(* IEC 61131-3 sources: Lasal-MCP/examples/SampleSource/5_ClassInputOutputSolution/Stations/MachineControl/MachineControl/Class/AlarmStation, 1 file *)

(* ---- AlarmStation.st ---- *)
(*!
<Class
	Name               = "AlarmStation"
	Revision           = "1.2"
	RealtimeTask       = "false"
	CyclicTask         = "false"
	BackgroundTask     = "false"
	Sigmatek           = "true"
	OSInterface        = "false"
	HighPriority       = "false"
	Automatic          = "false"
	UpdateMode         = "Prescan"
	SharedCommandTable = "true"
	Objectsize         = "(586,120)"
	Comment            = "Class collected number of active op-mode alarms and delivers this informations to the class AlarmBufferBase.">
	<Channels>
		<Server Name="ClassSvr" Visualized="false" Initialize="false" WriteProtected="true" Retentive="false"/>
		<Client Name="Active" Required="false" Internal="false"/>
		<Client Name="AlarmInfo" Required="false" Internal="false"/>
		<Client Name="coAlarmBufferBase" Required="true" Internal="false"/>
		<Client Name="GroupAutomatic" Required="false" Internal="false"/>
		<Client Name="GroupError" Required="false" Internal="false"/>
		<Client Name="GroupHoming" Required="false" Internal="false"/>
		<Client Name="GroupInit" Required="false" Internal="false"/>
		<Client Name="GroupManual" Required="false" Internal="false"/>
		<Client Name="GroupSemiAuto" Required="false" Internal="false"/>
		<Client Name="GroupSetup" Required="false" Internal="false"/>
		<Client Name="GroupStop" Required="false" Internal="false"/>
	</Channels>
	<RevDoku>
		<Owner Company="Sigmatek" Author="ObeChr"/>
		<Dokumentation Revision="1.2" Date="2017-07-26" Author="KruAle" Company="Sigmatek" Description="Added client to deactivate class if station is not available."/>
		<Dokumentation Revision="1.1" Date="2016-08-09" Author="ObeChr" Company="Sigmatek" Description="Added client to get AlarmInfo from other stations."/>
		<Dokumentation Revision="1.0" Date="2016-03-23" Author="ObeChr" Company="Sigmatek" Description="First library version."/>
	</RevDoku>
</Class>
*)
AlarmStation : CLASS
  //Servers:
	ClassSvr 	: SvrChCmd_DINT;
  //Clients:
	coAlarmBufferBase 	: CltChCmd_AlarmBufferBase;
	Active 	: CltCh_DINT;
	GroupInit 	: CltCh_UDINT;
	GroupHoming 	: CltCh_UDINT;
	GroupStop 	: CltCh_UDINT;
	GroupSetup 	: CltCh_UDINT;
	GroupManual 	: CltCh_UDINT;
	GroupSemiAuto 	: CltCh_UDINT;
	GroupAutomatic 	: CltCh_UDINT;
	GroupError 	: CltCh_UDINT;
	AlarmInfo 	: CltCh_BDINT;
  //Variables:
  //Functions:

	FUNCTION VIRTUAL GLOBAL Init;

	FUNCTION GLOBAL GetAlarms
		VAR_INPUT
			pAlarms 	: ^AlarmBufferBase::t_s_OPMode;
			pAlarmInfo 	: ^BDINT;
		END_VAR
		VAR_OUTPUT
			bSuccessful 	: BOOL;
		END_VAR;
  //Tables:
	FUNCTION @STD
		VAR_OUTPUT
			ret_code	: CONFSTATES;
		END_VAR;
	FUNCTION GLOBAL TAB @CT_;
END_CLASS;

#pragma usingLtd AlarmBufferBase

FUNCTION VIRTUAL GLOBAL AlarmStation::Init

  // last init-run
  if _FirstScan then

    // Login at AlarmBufferBase
    if coAlarmBufferBase.LoginAlarmClient(pThis := this) = false then
      TRACE_ERR("AlarmStation::Init(): login at AlarmBufferBase failed");
    end_if;

  end_if;

END_FUNCTION

FUNCTION GLOBAL AlarmStation::GetAlarms
	VAR_INPUT
		pAlarms 	: ^AlarmBufferBase::t_s_OPMode;
		pAlarmInfo 	: ^BDINT;
	END_VAR
	VAR_OUTPUT
		bSuccessful 	: BOOL;
	END_VAR

  // check input parameter
  if pAlarms = NIL | pAlarmInfo = NIL then
    bSuccessful := false;
    return;
  end_if;

  // check if station is active
  Active := Active.Read();
  if Active then

    // read client
    GroupInit       := GroupInit.Read();
    GroupHoming     := GroupHoming.Read();
    GroupStop       := GroupStop.Read();
    GroupSetup      := GroupSetup.Read();
    GroupManual     := GroupManual.Read();
    GroupSemiAuto   := GroupSemiAuto.Read();
    GroupAutomatic  := GroupAutomatic.Read();
    GroupError      := GroupError.Read();
    AlarmInfo       := AlarmInfo.Read();

  else
    GroupInit       := 0;
    GroupHoming     := 0;
    GroupStop       := 0;
    GroupSetup      := 0;
    GroupManual     := 0;
    GroupSemiAuto   := 0;
    GroupAutomatic  := 0;
    GroupError      := 0;
    AlarmInfo       := 0;
  end_if;

  // store opmode informations
  pAlarms^.udOPModeInit       := GroupInit;
  pAlarms^.udOPModeHoming     := GroupHoming;
  pAlarms^.udOPModeStop       := GroupStop;
  pAlarms^.udOPModeSetup      := GroupSetup;
  pAlarms^.udOPModeManual     := GroupManual;
  pAlarms^.udOPModeSemiAuto   := GroupSemiAuto;
  pAlarms^.udOPModeAutomatic  := GroupAutomatic;
  pAlarms^.udOPModeError      := GroupError;

  // store alarminfo
  pAlarmInfo^ := AlarmInfo;

  // set returncode
  bSuccessful := true;

END_FUNCTION
